TYPE "FRK_ProfileOwned_DeclarationUnit"
VERSION : 0.1
   STRUCT
      Book { ExternalAccessible := 'False'; ExternalVisible := 'False'; ExternalWritable := 'False'} : "FRK_ProfileBook";
      Steps { ExternalAccessible := 'False'; ExternalVisible := 'False'; ExternalWritable := 'False'} : Array[1..4] of "ST_StepTiming";
      LastSteps { ExternalAccessible := 'False'; ExternalVisible := 'False'; ExternalWritable := 'False'} : Array[1..4] of "ST_StepTiming";
      Stats { ExternalAccessible := 'False'; ExternalVisible := 'False'; ExternalWritable := 'False'} : Array[1..4] of "ST_TimingRow";
      History { ExternalAccessible := 'False'; ExternalVisible := 'False'; ExternalWritable := 'False'} : Array[1..60] of "ST_CycleSummary";
   END_STRUCT;

END_TYPE

